(* IEC 61131-3 sources: ia2/library/process-control/pous, 45 files *)

(* ---- fb_alarm_dev.st ---- *)
(*
  FB_ALARM_DEV — deviation alarm (pv over/under deviation from sp), deadband + delay + acknowledge latch.

  ~ Deviation alarm (over/under deviation), standard for loop monitoring.

  Purpose: loop-performance monitoring: alarm on a control deviation that persistently
  exceeds its limit (a stuck valve, an abrupt load change, lost tuning, a failed actuator).
  Behavior (follows the FB_ALARM_HL deadband+delay+latch pattern):
    dev := pv - sp.
    Over deviation:  dev > dev_h sets; dev < dev_h - deadband resets.
    Under deviation: dev < -dev_l sets; dev > -dev_l + deadband resets (dev_l supplied positive).
    Each trips after persisting for delay_s; output = trip OR (latched AND NOT ack)
    -- while the condition exists the alarm stays on, after it clears it is held until acknowledged.

  Inputs:
    pv       REAL  process value
    sp       REAL  setpoint (feed the same sp source as FB_PID; if the PID uses sp_rate,
                   prefer feeding the actual working sp after the ramp)
    dev_h    REAL  over-deviation limit (allowed amount pv may exceed sp)
    dev_l    REAL  under-deviation limit (allowed amount pv may fall below sp, supplied positive)
    deadband REAL  deadband (hysteresis, engineering units)
    delay_s  REAL  alarm delay s (0 = immediate)
    dt_s     REAL  sample period s
    ack      BOOL  acknowledge (level-active)
  Outputs:
    h_alm   BOOL  over-deviation alarm (latched)
    l_alm   BOOL  under-deviation alarm (latched)
    any_alm BOOL  any deviation alarm
*)
FUNCTION_BLOCK FB_ALARM_DEV
  VAR_INPUT
    pv       : REAL;
    sp       : REAL;
    dev_h    : REAL := 10.0;
    dev_l    : REAL := 10.0;
    deadband : REAL := 0.0;
    delay_s  : REAL := 0.0;
    dt_s     : REAL := 0.1;
    ack      : BOOL := FALSE;
  END_VAR
  VAR_OUTPUT
    h_alm   : BOOL;
    l_alm   : BOOL;
    any_alm : BOOL;
  END_VAR
  VAR
    dv     : REAL; (* pv - sp *)
    h_cond : BOOL;
    l_cond : BOOL;
    h_t    : REAL; (* delay accumulator, manual timing in place of TON *)
    l_t    : REAL;
    h_trip : BOOL;
    l_trip : BOOL;
  END_VAR

  dv := pv - sp;

  (* ---- Over deviation ---- *)
  IF dv > dev_h THEN
    h_cond := TRUE;
  ELSIF dv < dev_h - deadband THEN
    h_cond := FALSE;
  END_IF;
  IF h_cond THEN
    h_t := h_t + dt_s;
  ELSE
    h_t := 0.0;
  END_IF;
  h_trip := h_cond AND (h_t >= delay_s);
  h_alm  := h_trip OR (h_alm AND NOT ack);

  (* ---- Under deviation ---- *)
  IF dv < 0.0 - dev_l THEN
    l_cond := TRUE;
  ELSIF dv > 0.0 - dev_l + deadband THEN
    l_cond := FALSE;
  END_IF;
  IF l_cond THEN
    l_t := l_t + dt_s;
  ELSE
    l_t := 0.0;
  END_IF;
  l_trip := l_cond AND (l_t >= delay_s);
  l_alm  := l_trip OR (l_alm AND NOT ack);

  any_alm := h_alm OR l_alm;
END_FUNCTION_BLOCK

(* ---- fb_alarm_hl.st ---- *)
(*
  FB_ALARM_HL — four-level high/low alarm (H/L/HH/LL) with deadband, delay and simplified ISA-18.2 acknowledge latch.

  Purpose: high/low/high-high/low-low alarms for analog values such as level/temperature/pressure.
  Example: a vessel level LT alarm, with HH interlocking the feed shutdown.

  Behavior (same for each level, independently timed):
    1) Raw limit decision (with deadband hysteresis):
       High type: pv > sp sets; pv < sp - deadband resets.
       Low type:  pv < sp sets; pv > sp + deadband resets.
    2) Delay: the limit condition must persist for delay_s before tripping (internally
       timed by manual dt_s accumulation, not a TON instance, for easy offline testing
       and portability).
    3) Latch (simplified ISA-18.2): alarm output = trip condition OR (latched AND NOT ack).
       That is, while the condition exists the alarm stays on; after the condition
       clears it is held until ack acknowledges and clears it.

  Inputs:
    pv        REAL  process value
    h_sp      REAL  high alarm setpoint
    l_sp      REAL  low alarm setpoint
    hh_sp     REAL  high-high alarm setpoint
    ll_sp     REAL  low-low alarm setpoint
    deadband  REAL  deadband (hysteresis, engineering units)
    delay_s   REAL  alarm delay s (0 = immediate)
    dt_s      REAL  sample period s
    ack       BOOL  acknowledge (level-active)
  Outputs:
    h_alm / l_alm / hh_alm / ll_alm  BOOL  latched alarm outputs
    any_alm                          BOOL  any alarm
    h_cond / l_cond / hh_cond / ll_cond BOOL raw limit flags (with deadband, undelayed, unlatched)
*)
FUNCTION_BLOCK FB_ALARM_HL
  VAR_INPUT
    pv       : REAL;
    h_sp     : REAL := 80.0;
    l_sp     : REAL := 20.0;
    hh_sp    : REAL := 90.0;
    ll_sp    : REAL := 10.0;
    deadband : REAL := 0.0;
    delay_s  : REAL := 0.0;
    dt_s     : REAL := 0.1;
    ack      : BOOL := FALSE;
  END_VAR
  VAR_OUTPUT
    h_alm   : BOOL;
    l_alm   : BOOL;
    hh_alm  : BOOL;
    ll_alm  : BOOL;
    any_alm : BOOL;
    h_cond  : BOOL;
    l_cond  : BOOL;
    hh_cond : BOOL;
    ll_cond : BOOL;
  END_VAR
  VAR
    h_t     : REAL; (* per-level delay accumulator, manual timing in place of TON *)
    l_t     : REAL;
    hh_t    : REAL;
    ll_t    : REAL;
    h_trip  : BOOL;
    l_trip  : BOOL;
    hh_trip : BOOL;
    ll_trip : BOOL;
  END_VAR

  (* ---- High alarm H ---- *)
  IF pv > h_sp THEN
    h_cond := TRUE;
  ELSIF pv < h_sp - deadband THEN
    h_cond := FALSE;
  END_IF;
  IF h_cond THEN
    h_t := h_t + dt_s;
  ELSE
    h_t := 0.0;
  END_IF;
  h_trip := h_cond AND (h_t >= delay_s);
  h_alm  := h_trip OR (h_alm AND NOT ack);

  (* ---- Low alarm L ---- *)
  IF pv < l_sp THEN
    l_cond := TRUE;
  ELSIF pv > l_sp + deadband THEN
    l_cond := FALSE;
  END_IF;
  IF l_cond THEN
    l_t := l_t + dt_s;
  ELSE
    l_t := 0.0;
  END_IF;
  l_trip := l_cond AND (l_t >= delay_s);
  l_alm  := l_trip OR (l_alm AND NOT ack);

  (* ---- High-high alarm HH ---- *)
  IF pv > hh_sp THEN
    hh_cond := TRUE;
  ELSIF pv < hh_sp - deadband THEN
    hh_cond := FALSE;
  END_IF;
  IF hh_cond THEN
    hh_t := hh_t + dt_s;
  ELSE
    hh_t := 0.0;
  END_IF;
  hh_trip := hh_cond AND (hh_t >= delay_s);
  hh_alm  := hh_trip OR (hh_alm AND NOT ack);

  (* ---- Low-low alarm LL ---- *)
  IF pv < ll_sp THEN
    ll_cond := TRUE;
  ELSIF pv > ll_sp + deadband THEN
    ll_cond := FALSE;
  END_IF;
  IF ll_cond THEN
    ll_t := ll_t + dt_s;
  ELSE
    ll_t := 0.0;
  END_IF;
  ll_trip := ll_cond AND (ll_t >= delay_s);
  ll_alm  := ll_trip OR (ll_alm AND NOT ack);

  any_alm := h_alm OR l_alm OR hh_alm OR ll_alm;
END_FUNCTION_BLOCK

(* ---- fb_alarm_roc.st ---- *)
(*
  FB_ALARM_ROC — rate-of-change alarm, with derivative filtering, delay and acknowledge latch.

  ~ Rate-of-change alarm, with the derivative denoised by a first-order filter.

  Purpose: monitoring abnormal rates of change such as temperature runaway, abrupt
  pressure change, level collapse (leak/pipe break).
  Behavior:
    Raw derivative raw_roc := (pv - pv_prev) / dt_s;
    roc is raw_roc through an internal PT1 filter (time constant fixed at 3*dt_s,
    settling in about 4 scans) -- a single-scan difference is extremely sensitive to
    quantization/noise and will false-alarm without filtering; for stronger denoising
    put FB_LAG ahead of pv.
    |roc| > roc_limit trips after persisting for delay_s; latched until ack (same as the
    FB_ALARM_HL pattern: while the condition exists the alarm stays on, after it clears
    it is held until acknowledged).
    roc_limit <= 0 -> monitoring disabled (trip condition always FALSE; a latched output
    still needs ack to clear).
    The first scan only aligns pv_prev and does not evaluate the alarm (avoiding a
    spurious startup derivative); dt_s <= 0 -> hold.

  Inputs:
    pv        REAL  process value
    roc_limit REAL  rate-of-change limit |units|/s (bidirectional)
    delay_s   REAL  alarm delay s (0 = immediate)
    dt_s      REAL  sample period s
    ack       BOOL  acknowledge (level-active)
  Outputs:
    alm BOOL  rate-of-change alarm (latched)
    roc REAL  filtered rate of change units/s (signed, usable for trend display)
*)
FUNCTION_BLOCK FB_ALARM_ROC
  VAR_INPUT
    pv        : REAL;
    roc_limit : REAL := 10.0;
    delay_s   : REAL := 0.0;
    dt_s      : REAL := 0.1;
    ack       : BOOL := FALSE;
  END_VAR
  VAR_OUTPUT
    alm : BOOL;
    roc : REAL;
  END_VAR
  VAR
    pv_prev   : REAL;
    raw_roc   : REAL;
    t_f       : REAL; (* derivative filter time constant = 3*dt_s *)
    cond      : BOOL;
    trip      : BOOL;
    alm_t     : REAL; (* delay accumulator *)
    init_done : BOOL;
  END_VAR

  IF dt_s <= 0.0 THEN
    RETURN; (* hold *)
  END_IF;

  IF NOT init_done THEN
    pv_prev := pv; (* first-scan alignment, no alarm evaluation *)
    roc := 0.0;
    init_done := TRUE;
    RETURN;
  END_IF;

  raw_roc := (pv - pv_prev) / dt_s;
  pv_prev := pv;

  (* Internal PT1 denoising: t_f = 3*dt_s fixed (absorbs 1/4 of the new value each scan) *)
  t_f := 3.0 * dt_s;
  roc := roc + dt_s / (t_f + dt_s) * (raw_roc - roc);

  cond := FALSE;
  IF roc_limit > 0.0 THEN
    IF roc > roc_limit OR roc < 0.0 - roc_limit THEN
      cond := TRUE;
    END_IF;
  END_IF;

  IF cond THEN
    alm_t := alm_t + dt_s;
  ELSE
    alm_t := 0.0;
  END_IF;
  trip := cond AND (alm_t >= delay_s);
  alm := trip OR (alm AND NOT ack);
END_FUNCTION_BLOCK

(* ---- fb_alt2.st ---- *)
(*
  FB_ALT2 — dual-valve (dual-device) timed rotator, with two external permissives.

  Purpose: two diverter valves / two pumps rotating on a fixed period for wear balancing.
  Example: dual-permissive diverting with an iron remover + a packing scale:
  permissive1 (iron remover running) or permissive2 (packing scale ready) lost ->
  both valves close at once; after the permissives recover, rotation continues by its
  timer (the rotation selection is held, the timer is cleared and restarts).

  Behavior:
    ok := enable AND permissive1 AND permissive2.
    NOT ok: q1 := FALSE, q2 := FALSE, rotation timer cleared (the selection bit is held,
    and after recovery continues from the last selected channel).
    ok: the timer accumulates by dt_s manually, and at swap_period_s the selection
    switches and the timer clears; q1/q2 output the currently selected channel mutually
    exclusively. swap_period_s <= 0 means no rotation (hold the current channel).

  Inputs:
    enable        BOOL  enable
    swap_period_s REAL  rotation period s
    dt_s          REAL  sample period s
    permissive1   BOOL  external permissive 1 (e.g. iron remover running)
    permissive2   BOOL  external permissive 2 (e.g. packing scale ready)
  Outputs:
    q1 BOOL  valve 1 output
    q2 BOOL  valve 2 output (mutually exclusive with q1; both FALSE when a permissive is lost)
*)
FUNCTION_BLOCK FB_ALT2
  VAR_INPUT
    enable        : BOOL;
    swap_period_s : REAL := 300.0;
    dt_s          : REAL := 0.1;
    permissive1   : BOOL := TRUE;
    permissive2   : BOOL := TRUE;
  END_VAR
  VAR_OUTPUT
    q1 : BOOL;
    q2 : BOOL;
  END_VAR
  VAR
    ok    : BOOL;
    sel2  : BOOL; (* FALSE selects valve 1 / TRUE selects valve 2, held while disabled *)
    run_t : REAL; (* this channel's elapsed run time s, manual timing *)
  END_VAR

  ok := enable AND permissive1 AND permissive2;

  IF NOT ok THEN
    (* Any permissive lost: both valves close, timer cleared, selection held *)
    q1    := FALSE;
    q2    := FALSE;
    run_t := 0.0;
    RETURN;
  END_IF;

  IF dt_s > 0.0 THEN
    run_t := run_t + dt_s;
  END_IF;
  IF swap_period_s > 0.0 AND run_t >= swap_period_s THEN
    run_t := 0.0;
    sel2  := NOT sel2;
  END_IF;

  q1 := NOT sel2;
  q2 := sel2;
END_FUNCTION_BLOCK

(* ---- fb_avg_time.st ---- *)
(*
  FB_AVG_TIME — tumbling-window time average.

  ~ Standard time-average block, the customary form for DCS reporting / steady-quantity monitoring.

  Purpose: full-window averages for reports (e.g. per-minute average flow), noise-robust
  readings of slowly varying quantities, drift monitoring by comparison against the
  instantaneous value.
  Behavior:
    Within the window, sum / count accumulate each scan; avg_run := sum / count is the
    running mean of the current window; when the window is full (accumulated time
    reaches window_s) avg_run is copied into avg, ready is set, and then the
    accumulators are cleared to start the next window (phase subtraction wraps so the
    long-term cadence does not drift).
    While the first window is not yet full, avg temporarily tracks avg_run (to avoid
    outputting 0 at startup) and ready = FALSE flags "not yet a complete-window result";
    after the first window completes ready stays TRUE and avg refreshes only on the
    window-full scan.
    reset level-active: clears the accumulators and ready, restarting the window.
    window_s <= 0 -> pass-through (avg := avg_run := u, ready := TRUE);
    dt_s <= 0 -> hold (no action).
    Note: this block is a tumbling window (one value per window), not a sliding window
    -- a true sliding window needs an array buffer (in this dialect an FB-scope array
    cannot be codegen'd, see README gotcha 7); for continuous "smoothed every scan"
    output, use FB_LAG exponential smoothing as an approximation.

  Inputs:
    u        REAL  input
    window_s REAL  averaging window length s (<= 0 pass-through)
    dt_s     REAL  sample period s
    reset    BOOL  reset (level-active: clear the window and restart)
  Outputs:
    avg     REAL  average of the previous complete window (tracks avg_run while the first window is incomplete)
    avg_run REAL  running mean of the current window
    ready   BOOL  first complete window has finished (avg is trustworthy)
*)
FUNCTION_BLOCK FB_AVG_TIME
  VAR_INPUT
    u        : REAL;
    window_s : REAL := 60.0;
    dt_s     : REAL := 0.1;
    reset    : BOOL := FALSE;
  END_VAR
  VAR_OUTPUT
    avg     : REAL;
    avg_run : REAL;
    ready   : BOOL;
  END_VAR
  VAR
    sum       : REAL; (* current-window accumulated sum *)
    count     : REAL; (* current-window sample count *)
    elapsed_s : REAL; (* current-window accumulated time, manual timing *)
  END_VAR

  IF reset THEN
    sum := 0.0;
    count := 0.0;
    elapsed_s := 0.0;
    avg := 0.0;
    avg_run := 0.0;
    ready := FALSE;
    RETURN;
  END_IF;

  IF window_s <= 0.0 THEN
    avg := u; (* invalid window length: pass-through *)
    avg_run := u;
    ready := TRUE;
    RETURN;
  END_IF;

  IF dt_s <= 0.0 THEN
    RETURN; (* invalid sample period: hold *)
  END_IF;

  sum := sum + u;
  count := count + 1.0;
  elapsed_s := elapsed_s + dt_s;
  avg_run := sum / count;

  IF elapsed_s >= window_s THEN
    (* Window full: copy the result, clear to start the next window (subtraction wrap keeps the long-term cadence) *)
    avg := avg_run;
    ready := TRUE;
    sum := 0.0;
    count := 0.0;
    elapsed_s := elapsed_s - window_s;
  ELSIF NOT ready THEN
    avg := avg_run; (* first window not yet full: avg tracks the running mean to avoid outputting 0 at startup *)
  END_IF;
END_FUNCTION_BLOCK

(* ---- fb_cascade.st ---- *)
(*
  FB_CASCADE — cascade coupling glue (master output -> slave SP mapping + non-cascade tracking back-calculation).

  ~ Standard cascade-coupling block (cascade SP coupling / master tracking
  back-calculation), the customary glue for cascade-loop configuration: only this one
  block sits between the two PIDs.

  Purpose: cascade-loop configuration (temperature master -> flow slave, and the like),
  mapping the master output 0..100% to the slave SP engineering span, and supplying the
  master a tracking value when not in cascade so that putting CAS into/out of service is
  bumpless.
  Behavior:
    CAS (cas_on = TRUE):
      slave_sp := sp_min + master_out / 100 * (sp_max - sp_min)
      master_track := FALSE (the master controls normally).
    Non-CAS:
      slave_sp := slave_sp_local (the operator's local SP given directly to the slave loop);
      master_track := TRUE, master_track_value :=
        (slave_sp_now - sp_min) / (sp_max - sp_min) * 100, clamped 0..100
      -- the master output is forced to "the equivalent percentage of the current slave
      SP", so on the scan that switches back to CAS slave_sp does not jump (bumpless transfer).
      Span not configured (|sp_max - sp_min| < 1E-6) -> tracking value takes 0 (divide-by-zero guard).
    The tracking value is computed every scan (independent of mode), so it is valid the
    instant CAS is removed.
    Pure combinational logic, no internal state.

  Wiring (cascading two FB_PID instances; slave_sp_now is fed the previous scan's working SP):
    casc(master_out := pid_master.out, cas_on := cas_enable,
         sp_min := 0.0, sp_max := 2000.0,
         slave_sp_local := op_sp, slave_sp_now := slave_sp_used);
    slave_sp_used := casc.slave_sp;
    pid_master(pv := temp_pv, sp := temp_sp, ..., dt_s := scan_s,
               track := casc.master_track,
               track_value := casc.master_track_value);
    pid_slave(pv := flow_pv, sp := slave_sp_used, ..., dt_s := scan_s);

  Inputs:
    master_out     REAL  master output 0..100 %
    cas_on         BOOL  cascade enabled (FALSE = slave uses local SP, master tracks)
    sp_min         REAL  slave SP span low (engineering units)
    sp_max         REAL  slave SP span high
    slave_sp_local REAL  slave-loop local SP when not in cascade
    slave_sp_now   REAL  slave-loop current working SP (feed the previous scan's slave_sp, for the tracking back-calculation)
  Outputs:
    slave_sp           REAL  slave-loop setpoint (to pid_slave.sp)
    master_track       BOOL  master tracking command (to pid_master.track)
    master_track_value REAL  master tracking value 0..100 % (to pid_master.track_value)
*)
FUNCTION_BLOCK FB_CASCADE
  VAR_INPUT
    master_out     : REAL;
    cas_on         : BOOL := FALSE;
    sp_min         : REAL := 0.0;
    sp_max         : REAL := 100.0;
    slave_sp_local : REAL := 0.0;
    slave_sp_now   : REAL := 0.0;
  END_VAR
  VAR_OUTPUT
    slave_sp           : REAL;
    master_track       : BOOL;
    master_track_value : REAL;
  END_VAR
  VAR
    span : REAL; (* slave-loop SP span width *)
  END_VAR

  span := sp_max - sp_min;

  (* Tracking value computed every scan: the equivalent percentage of the current slave SP (span not configured -> 0, divide-by-zero guard) *)
  IF (span < 0.000001) AND (span > -0.000001) THEN
    master_track_value := 0.0;
  ELSE
    master_track_value := (slave_sp_now - sp_min) / span * 100.0;
    IF master_track_value < 0.0 THEN
      master_track_value := 0.0;
    ELSIF master_track_value > 100.0 THEN
      master_track_value := 100.0;
    END_IF;
  END_IF;

  IF cas_on THEN
    slave_sp := sp_min + master_out / 100.0 * span;
    master_track := FALSE;
  ELSE
    slave_sp := slave_sp_local;
    master_track := TRUE;
  END_IF;
END_FUNCTION_BLOCK

(* ---- fb_char.st ---- *)
(*
  FB_CHAR — piecewise-linear signal characterization (linear interpolation, up to 8 points).

  ~ Piecewise-linear characterizer, the customary block for valve-characteristic linearization / nonlinear sensors.

  Purpose: valve-characteristic linearization (equal-percentage valve-opening
  compensation), nonlinear sensor calibration, level-to-volume conversion, and any
  monotonic piecewise-linear transform.

  Behavior:
    Take the first n points (x1,y1)..(xn,yn) (n clamped to 2..8); interpolate
    linearly when u falls in segment (xk, xk+1]; u <= x1 -> out := y1; u >= xn ->
    out := yn (clamped at both ends).
    Convention: x must be ascending (no hard check here; a degenerate non-ascending
    segment yields the right-end y).
    In this dialect an ARRAY in FUNCTION_BLOCK scope cannot be codegen'd (see the
    README dialect gotchas), so scalar point pairs x1..x8 / y1..y8 + n are used.

  Inputs:
    u          REAL  input
    n          INT   number of points in use 2..8 (auto-clamped)
    x1..x8     REAL  breakpoint x coordinates (ascending)
    y1..y8     REAL  breakpoint y coordinates
  Outputs:
    out        REAL  characterized output (clamped at both ends)
*)
FUNCTION_BLOCK FB_CHAR
  VAR_INPUT
    u  : REAL;
    n  : INT := 2;
    x1 : REAL := 0.0;
    y1 : REAL := 0.0;
    x2 : REAL := 100.0;
    y2 : REAL := 100.0;
    x3 : REAL := 0.0;
    y3 : REAL := 0.0;
    x4 : REAL := 0.0;
    y4 : REAL := 0.0;
    x5 : REAL := 0.0;
    y5 : REAL := 0.0;
    x6 : REAL := 0.0;
    y6 : REAL := 0.0;
    x7 : REAL := 0.0;
    y7 : REAL := 0.0;
    x8 : REAL := 0.0;
    y8 : REAL := 0.0;
  END_VAR
  VAR_OUTPUT
    out : REAL;
  END_VAR
  VAR
    nn    : INT;  (* clamped point count *)
    xa    : REAL; (* selected segment left end *)
    ya    : REAL;
    xb    : REAL; (* selected segment right end *)
    yb    : REAL;
    span  : REAL;
    found : BOOL;
  END_VAR

  nn := n;
  IF nn < 2 THEN
    nn := 2;
  ELSIF nn > 8 THEN
    nn := 8;
  END_IF;

  (* Low-end clamp *)
  IF u <= x1 THEN
    out := y1;
    RETURN;
  END_IF;

  (* Segment search: take the segment u falls into, (xk, xk+1]; only the first nn points are considered *)
  found := FALSE;
  IF u <= x2 THEN
    xa := x1; ya := y1; xb := x2; yb := y2; found := TRUE;
  ELSIF nn >= 3 AND u <= x3 THEN
    xa := x2; ya := y2; xb := x3; yb := y3; found := TRUE;
  ELSIF nn >= 4 AND u <= x4 THEN
    xa := x3; ya := y3; xb := x4; yb := y4; found := TRUE;
  ELSIF nn >= 5 AND u <= x5 THEN
    xa := x4; ya := y4; xb := x5; yb := y5; found := TRUE;
  ELSIF nn >= 6 AND u <= x6 THEN
    xa := x5; ya := y5; xb := x6; yb := y6; found := TRUE;
  ELSIF nn >= 7 AND u <= x7 THEN
    xa := x6; ya := y6; xb := x7; yb := y7; found := TRUE;
  ELSIF nn >= 8 AND u <= x8 THEN
    xa := x7; ya := y7; xb := x8; yb := y8; found := TRUE;
  END_IF;

  IF found THEN
    span := xb - xa;
    IF span > 0.0 THEN
      out := ya + (u - xa) * (yb - ya) / span;
    ELSE
      out := yb; (* degenerate segment (x not ascending): take the right end *)
    END_IF;
    RETURN;
  END_IF;

  (* High-end clamp: u greater than the nn-th point *)
  CASE nn OF
    3:
      out := y3;
    4:
      out := y4;
    5:
      out := y5;
    6:
      out := y6;
    7:
      out := y7;
    8:
      out := y8;
  ELSE
    out := y2;
  END_CASE;
END_FUNCTION_BLOCK

(* ---- fb_deadtime8.st ---- *)
(*
  FB_DEADTIME8 — dead time / transport delay, 8 scalar taps + linear interpolation.

  ~ Standard dead-time block (dead time / PTt / transport delay), the customary block
  for plant simulation and feedforward dynamic compensation (Smith-predictor-type structures).

  Purpose: plant simulation (in series with FB_LAG it forms a first-order-lag-plus-dead-time
  FOPDT plant), transport-delay matching in a feedforward path, time alignment of
  belt/pipe-conveying measurements.
  Behavior:
    Tap chain z1..z8 (z1 newest, z8 oldest), sampling interval = t_delay_s / 8:
    the phase phase_s accumulates by dt_s manually, and each time a sampling interval
    elapses the whole chain shifts once (z8<-z7<-...<-z1<-u); at most 8 shifts per scan
    (after 8 the whole chain has been filled by u, so the WHILE is bounded and
    scan-deterministic).
    The output interpolates linearly between the two oldest taps by the phase fraction:
      out := z8 + (z7 - z8) * phase_s / period_s
    -- a step input is traversed as a ramp over one sampling interval, so the output is
       continuous with no steps.
    Resolution = t_delay_s / 8: 8 taps is the compromise in an array-free dialect; the
    staircase/interpolation error of the delay time is about 1/8 of the delay --
    adequate for loop tuning; for finer resolution, put two of these blocks in series
    (each carrying half the delay).
    t_delay_s <= 0 -> pass-through (out := u), and the taps fill with u -- when the
    delay is put into service online it starts smoothly from the current value (bumpless).
    reset / first scan: all taps filled with u, out := u, phase cleared.
    dt_s <= 0 -> hold (no action).

  Inputs:
    u         REAL  input
    t_delay_s REAL  dead time s (<= 0 pass-through; changeable online, advances at the new interval)
    dt_s      REAL  sample period s
    reset     BOOL  reset (level-active: taps filled with u, output follows u)
  Outputs:
    out REAL  delayed output (linearly interpolated, continuous)
*)
FUNCTION_BLOCK FB_DEADTIME8
  VAR_INPUT
    u         : REAL;
    t_delay_s : REAL := 0.0;
    dt_s      : REAL := 0.1;
    reset     : BOOL := FALSE;
  END_VAR
  VAR_OUTPUT
    out : REAL;
  END_VAR
  VAR
    z1        : REAL; (* tap chain: z1 newest ... z8 oldest (scalar form for the array-free dialect) *)
    z2        : REAL;
    z3        : REAL;
    z4        : REAL;
    z5        : REAL;
    z6        : REAL;
    z7        : REAL;
    z8        : REAL;
    phase_s   : REAL; (* phase within the current sampling interval, manual timing *)
    period_s  : REAL; (* sampling interval = t_delay_s / 8 *)
    shifts    : REAL; (* shift count this scan (capped at 8: chain already saturated) *)
    init_done : BOOL; (* first-scan alignment flag *)
  END_VAR

  IF reset OR NOT init_done THEN
    z1 := u;
    z2 := u;
    z3 := u;
    z4 := u;
    z5 := u;
    z6 := u;
    z7 := u;
    z8 := u;
    phase_s := 0.0;
    out := u;
    init_done := TRUE;
    RETURN;
  END_IF;

  IF t_delay_s <= 0.0 THEN
    (* Pass-through; taps fill with u, so when the delay is put into service online it starts bumplessly from the current value *)
    z1 := u;
    z2 := u;
    z3 := u;
    z4 := u;
    z5 := u;
    z6 := u;
    z7 := u;
    z8 := u;
    phase_s := 0.0;
    out := u;
    RETURN;
  END_IF;

  IF dt_s <= 0.0 THEN
    RETURN; (* invalid sample period: hold *)
  END_IF;

  period_s := t_delay_s / 8.0;
  phase_s := phase_s + dt_s;

  (* Shift the whole chain once per elapsed sampling interval; capped at 8/scan (when
     dt_s spans several intervals, catch up; after 8 the chain is full of u and further
     shifts are meaningless) -- the WHILE is bounded *)
  shifts := 0.0;
  WHILE (phase_s >= period_s) AND (shifts < 8.0) DO
    z8 := z7;
    z7 := z6;
    z6 := z5;
    z5 := z4;
    z4 := z3;
    z3 := z2;
    z2 := z1;
    z1 := u;
    phase_s := phase_s - period_s;
    shifts := shifts + 1.0;
  END_WHILE;
  IF phase_s >= period_s THEN
    phase_s := 0.0; (* degenerate case dt_s >= t_delay_s: chain is already u, clear phase to prevent accumulation *)
  END_IF;

  (* Interpolate between the two oldest taps by phase fraction: at the shift instant frac=0 -> out=z8(old z7), continuous *)
  out := z8 + (z7 - z8) * phase_s / period_s;
END_FUNCTION_BLOCK

(* ---- fb_debounce.st ---- *)
(*
  FB_DEBOUNCE — discrete-input debounce (independent bidirectional confirmation delay).

  ~ Discrete-input debounce (on/off dual delay), standard for DI processing.

  Purpose: confirming chattering signals such as float level switches, limit switches,
  relay/contactor auxiliary contacts; can also debounce the run_fb/fault inputs of
  FB_DUTY2.
  Behavior:
    u continuously TRUE for t_on_s -> q := TRUE; u continuously FALSE for t_off_s ->
    q := FALSE; any reverse transition in between clears that direction's timer (restart).
    t = 0 means that direction takes effect immediately. The actual confirmation time
    rounds up to a dt_s scan.
    (Manual dt_s accumulation, equivalent to a TON on-confirm + off-confirm, offline-testable.)

  Inputs:
    u       BOOL  raw discrete input
    t_on_s  REAL  set confirmation time s (0 = immediate)
    t_off_s REAL  reset confirmation time s (0 = immediate)
    dt_s    REAL  sample period s
  Outputs:
    q       BOOL  debounced discrete output
*)
FUNCTION_BLOCK FB_DEBOUNCE
  VAR_INPUT
    u       : BOOL;
    t_on_s  : REAL := 0.1;
    t_off_s : REAL := 0.1;
    dt_s    : REAL := 0.1;
  END_VAR
  VAR_OUTPUT
    q : BOOL;
  END_VAR
  VAR
    on_t  : REAL; (* set-direction accumulator *)
    off_t : REAL; (* reset-direction accumulator *)
  END_VAR

  IF u THEN
    off_t := 0.0;
    IF NOT q THEN
      on_t := on_t + dt_s;
      IF on_t >= t_on_s THEN
        q := TRUE;
      END_IF;
    END_IF;
  ELSE
    on_t := 0.0;
    IF q THEN
      off_t := off_t + dt_s;
      IF off_t >= t_off_s THEN
        q := FALSE;
      END_IF;
    END_IF;
  END_IF;
END_FUNCTION_BLOCK

(* ---- fb_deriv.st ---- *)
(*
  FB_DERIV — filtered derivative (du/dt, filter first then difference).

  ~ Standard filtered-derivative block, a staple of every major platform's standard library.

  Purpose: quantifying trend (degC/s, %/s for display/feedforward/custom logic),
  derivative shaping in a feedforward path. Whenever you want "alarm on limit", use
  FB_ALARM_ROC directly (the same filter-difference core + delay/latch).
  Behavior:
    u first passes through an internal PT1 filter (time constant t_filt_s; <= 0 takes
    3*dt_s automatically, settling in about 4 scans), then a backward difference of
    the filtered value:
      u_f := u_f + dt_s / (t_f + dt_s) * (u - u_f)
      out := (u_f - u_f_prev) / dt_s
    A single-scan difference is extremely sensitive to quantization/noise and must be
    filtered, or the output is all spikes -- for stronger noise rejection, increase
    t_filt_s or put FB_LAG ahead of u.
    reset / first scan: the filter state aligns to u, out := 0 (no spurious startup derivative).
    dt_s <= 0 -> hold (no action).

  Inputs:
    u        REAL  input
    t_filt_s REAL  derivative pre-filter time constant s (<= 0 = auto 3*dt_s)
    dt_s     REAL  sample period s
    reset    BOOL  reset/align (level-active: filter state follows u, out cleared)
  Outputs:
    out REAL  filtered rate of change units/s (signed)
*)
FUNCTION_BLOCK FB_DERIV
  VAR_INPUT
    u        : REAL;
    t_filt_s : REAL := 0.0;
    dt_s     : REAL := 0.1;
    reset    : BOOL := FALSE;
  END_VAR
  VAR_OUTPUT
    out : REAL;
  END_VAR
  VAR
    u_f       : REAL; (* PT1-filtered input *)
    u_f_prev  : REAL; (* previous-scan filtered value, for the backward difference *)
    t_f       : REAL; (* filter time constant actually used *)
    init_done : BOOL; (* first-scan alignment flag *)
  END_VAR

  IF dt_s <= 0.0 THEN
    RETURN; (* invalid sample period: hold *)
  END_IF;

  IF reset OR NOT init_done THEN
    u_f := u; (* align the filter state, no spurious startup derivative *)
    u_f_prev := u;
    out := 0.0;
    init_done := TRUE;
    RETURN;
  END_IF;

  t_f := t_filt_s;
  IF t_f <= 0.0 THEN
    t_f := 3.0 * dt_s; (* auto: the minimum noise rejection that settles in about 4 scans *)
  END_IF;

  u_f := u_f + dt_s / (t_f + dt_s) * (u - u_f);
  out := (u_f - u_f_prev) / dt_s;
  u_f_prev := u_f;
END_FUNCTION_BLOCK

(* ---- fb_dose.st ---- *)
(*
  FB_DOSE — batch dosing / batch feeding (coarse/fine two stages + in-flight compensation).

  ~ Standard dosing block (dosing / batch weighing, coarse-fine two-speed feeding +
  early in-flight cutoff), the customary block for batch-scale / batch-feed control.

  Purpose: dosing material from a silo into a weigh hopper / reactor: coarse feed
  approaches the target quickly, fine feed trims, the fine valve closes early by the
  in-flight amount (the material still in flight after the valve closes), and after
  settling the completion and overshoot are reported. The flow input may come from a
  weight derivative or a flowmeter.

  Behavior:
    start rising edge (when idle, not complete, and abort not pressed) begins a new
    batch: qty cleared, enter the feed stage. During feeding/settling, accumulate
    qty := qty + flow * dt_s (flow <= 0 not counted, one of the criteria for material
    fully landed).
      Coarse stage: qty < target - fine_qty -> q_coarse = TRUE (both coarse and fine valves open);
      Fine stage: qty < target - inflight -> q_fine = TRUE; at the point, close the fine
      valve (the in-flight reserve inflight is the in-flight amount held back) and enter
      the settling stage.
      Settling stage: wait for flow <= 0 or a fixed 2 s (whichever first) -> done := TRUE,
      overshoot := qty - target (the actual overshoot once the in-flight material has landed).
    abort level-active: stop both valves immediately, exit feeding/settling, qty
    retained (for stocktaking), done not set.
    After done, start has no effect; reset (level-active) is required to clear
    qty/done/overshoot and begin the next batch.
    Assumes fine_qty >= inflight >= 0 (coarse valve closes first, fine valve closes after);
    dribble after done is no longer counted into qty.
    dt_s <= 0 -> hold this scan, no action (command edges still remembered).

  Inputs:
    start    BOOL  start (rising edge begins a new batch)
    abort    BOOL  abort (level-active: stop valves, retain quantity)
    flow     REAL  instantaneous flow units/s (weight derivative or flowmeter)
    target   REAL  target quantity (same unit as the flow integral)
    fine_qty REAL  fine-feed-stage quantity (close the coarse valve with this much remaining)
    inflight REAL  in-flight amount (close the fine valve with this much remaining)
    dt_s     REAL  sample period s
    reset    BOOL  batch reset (level-active: clear qty/done/overshoot)
  Outputs:
    q_coarse  BOOL  coarse-feed valve
    q_fine    BOOL  fine-feed valve
    qty       REAL  this batch's accumulated quantity
    done      BOOL  this batch complete (set after settling, held until reset)
    overshoot REAL  actual - target after completion (basis for tuning the in-flight amount)
*)
FUNCTION_BLOCK FB_DOSE
  VAR_INPUT
    start    : BOOL;
    abort    : BOOL;
    flow     : REAL;
    target   : REAL := 100.0;
    fine_qty : REAL := 10.0;
    inflight : REAL := 0.0;
    dt_s     : REAL := 0.1;
    reset    : BOOL;
  END_VAR
  VAR_OUTPUT
    q_coarse  : BOOL;
    q_fine    : BOOL;
    qty       : REAL;
    done      : BOOL;
    overshoot : REAL;
  END_VAR
  VAR
    dosing     : BOOL; (* feed stage (coarse/fine) *)
    settling   : BOOL; (* settling-wait stage *)
    settle_t   : REAL; (* settling timer s *)
    prev_start : BOOL; (* start rising-edge memory *)
  END_VAR

  IF reset THEN
    dosing     := FALSE;
    settling   := FALSE;
    settle_t   := 0.0;
    qty        := 0.0;
    done       := FALSE;
    overshoot  := 0.0;
    q_coarse   := FALSE;
    q_fine     := FALSE;
    prev_start := start;
    RETURN;
  END_IF;

  IF abort THEN
    (* Abort: stop valves and exit the stage, qty retained, done not set *)
    dosing   := FALSE;
    settling := FALSE;
    q_coarse := FALSE;
    q_fine   := FALSE;
  END_IF;

  (* start rising edge, idle and not complete -> begin a new batch *)
  IF start AND NOT prev_start AND NOT abort
     AND NOT dosing AND NOT settling AND NOT done THEN
    dosing    := TRUE;
    qty       := 0.0;
    overshoot := 0.0;
    settle_t  := 0.0;
  END_IF;
  prev_start := start;

  IF dt_s <= 0.0 THEN
    RETURN; (* invalid sample period: hold *)
  END_IF;

  (* Accumulate flow during feeding/settling (negative flow not counted) *)
  IF (dosing OR settling) AND flow > 0.0 THEN
    qty := qty + flow * dt_s;
  END_IF;

  IF dosing THEN
    q_coarse := qty < target - fine_qty;
    q_fine   := qty < target - inflight;
    IF NOT q_fine THEN
      (* At the in-flight reserve point: close the fine valve and enter the settling stage *)
      q_coarse := FALSE;
      dosing   := FALSE;
      settling := TRUE;
      settle_t := 0.0;
    END_IF;
  END_IF;

  IF settling THEN
    settle_t := settle_t + dt_s;
    IF flow <= 0.0 OR settle_t >= 2.0 THEN
      settling  := FALSE;
      done      := TRUE;
      overshoot := qty - target;
    END_IF;
  END_IF;
END_FUNCTION_BLOCK

(* ---- fb_duty2.st ---- *)
(*
  FB_DUTY2 — dual-pump duty/standby rotation control.

  ~ Dual-pump duty/standby rotation: select the duty pump by start sequence or run-hour
  balancing, with immediate takeover on fault.

  Purpose: two pumps in a duty/standby arrangement: select the duty pump by rotating
  each start or by balancing accumulated run hours; on a duty-pump fault the standby
  takes over immediately; on a dual fault both stop.
  Behavior (scan-deterministic: no internal timing, only edge memory):
    A demand rising edge selects this round's duty pump, by priority:
      1) exactly one is already running (run_fb TRUE on one side) -> adopt it as duty
         directly (bumpless takeover, avoiding stopping it to start the standby);
      2) alt_mode = 1 -> the lower accumulated hours is duty (hours_a/b fed from two FB_RUNTIME);
      3) alt_mode = 0 (default) -> toggle from the current duty position (including the
         state after a fault takeover, giving natural wear balancing).
    While demand persists: a duty-pump fault with the other healthy -> duty switches
    immediately (takeover); a commanded pump that faults gets no command; a dual fault
    -> both cmd FALSE (the duty selection is held).
    demand withdrawn -> both cmd FALSE.
    Wiring suggestion: feed fault_x from FB_MOTOR's fault or the electrical protection
    relay; feed run_fb_x from the run feedback (debounce a chattering contact with
    FB_DEBOUNCE); leave feedback-timeout fault decision to FB_MOTOR, this block does not
    duplicate the timing.

  Inputs:
    demand   BOOL  system needs a pump (level)
    alt_mode INT   0 = rotate each start / 1 = run-hour balancing
    run_fb_a BOOL  pump A run feedback
    run_fb_b BOOL  pump B run feedback
    fault_a  BOOL  pump A fault
    fault_b  BOOL  pump B fault
    hours_a  REAL  pump A accumulated hours (used by alt_mode=1, fed from FB_RUNTIME.hours)
    hours_b  REAL  pump B accumulated hours (used by alt_mode=1)
    dt_s     REAL  sample period s (this block does not currently time; kept for a uniform library interface)
  Outputs:
    cmd_a     BOOL  pump A start command
    cmd_b     BOOL  pump B start command
    duty_is_a BOOL  the current duty pump is A
*)
FUNCTION_BLOCK FB_DUTY2
  VAR_INPUT
    demand   : BOOL;
    alt_mode : INT := 0;
    run_fb_a : BOOL := FALSE;
    run_fb_b : BOOL := FALSE;
    fault_a  : BOOL := FALSE;
    fault_b  : BOOL := FALSE;
    hours_a  : REAL := 0.0;
    hours_b  : REAL := 0.0;
    dt_s     : REAL := 0.1;
  END_VAR
  VAR_OUTPUT
    cmd_a     : BOOL;
    cmd_b     : BOOL;
    duty_is_a : BOOL;
  END_VAR
  VAR
    prev_demand : BOOL; (* rising-edge memory *)
    rising      : BOOL;
  END_VAR

  rising := demand AND NOT prev_demand;
  prev_demand := demand;

  IF rising THEN
    IF run_fb_a AND NOT run_fb_b THEN
      duty_is_a := TRUE;  (* the already-running pump becomes duty directly, bumpless takeover *)
    ELSIF run_fb_b AND NOT run_fb_a THEN
      duty_is_a := FALSE;
    ELSIF alt_mode = 1 THEN
      duty_is_a := hours_a <= hours_b; (* hour balancing: the lower is duty *)
    ELSE
      duty_is_a := NOT duty_is_a; (* rotate each start (initial FALSE -> first start selects A) *)
    END_IF;
  END_IF;

  IF demand THEN
    (* Fault takeover: duty faults and the other is healthy -> duty switches immediately *)
    IF duty_is_a AND fault_a AND NOT fault_b THEN
      duty_is_a := FALSE;
    ELSIF NOT duty_is_a AND fault_b AND NOT fault_a THEN
      duty_is_a := TRUE;
    END_IF;
    cmd_a := duty_is_a AND NOT fault_a;
    cmd_b := NOT duty_is_a AND NOT fault_b;
  ELSE
    cmd_a := FALSE;
    cmd_b := FALSE;
  END_IF;
END_FUNCTION_BLOCK

(* ---- fb_flow_comp.st ---- *)
(*
  FB_FLOW_COMP — gas-flow pressure/temperature compensation (ideal-gas approximation).

  ~ Standard pressure/temperature compensation block for gas flow, the customary
  block for correcting gas flow to standard / design conditions.

  Purpose: correct gas flow to reference (design) conditions using operating
  pressure/temperature: reading correction for a DP flowmeter calibrated at design
  conditions when operation departs from the design point, and correction of
  volumetric flow to standard conditions. Compensation ratio:
    ratio := (p_abs / p_ref) * (t_ref_k / t_k)   -- density ratio (ideal gas)
    p_abs := p_gauge_kpa + atm_kpa (gauge -> absolute)
    t_k   := t_c + 273.15
  Behavior (mode selects the flowmeter type):
    mode = 0 (square-root DP flowmeter, the flow signal after DP square-root extraction):
      q_comp := q_raw * SQRT(ratio)
      -- DP flow is proportional to SQRT(density), so a density departure from the
         design value is corrected via the square root.
    mode = 1 (linear volumetric, operating volumetric flow corrected to reference conditions):
      q_comp := q_raw * ratio
    Guard: t_k <= 0, t_ref_k <= 0, p_ref_kpa_abs <= 0 or p_abs <= 0
    (invalid measurement/configuration) -> q_comp := q_raw pass-through.
    Pure combinational logic, no internal state.
    Scope note: ideal-gas approximation (no compressibility-factor or humidity
    correction); custody-transfer-grade full-specification energy-metering standard
    algorithms are outside this block's scope.
    Reference conditions default to p_ref = 201.325 kPa(a) (i.e. 100 kPa gauge +
    standard atmosphere), t_ref = 20 degC -- set per the flowmeter design datasheet.

  Inputs:
    q_raw         REAL  raw flow (operating reading)
    p_gauge_kpa   REAL  operating gauge pressure kPa(g)
    t_c           REAL  operating temperature degC
    p_ref_kpa_abs REAL  reference absolute pressure kPa(a) (design condition)
    t_ref_c       REAL  reference temperature degC (design condition)
    atm_kpa       REAL  local atmospheric pressure kPa (gauge -> absolute conversion)
    mode          REAL  0 = square-root DP (multiply by SQRT(ratio)) /
                        1 = linear volumetric (multiply by ratio)
  Outputs:
    q_comp REAL  compensated flow
*)
FUNCTION_BLOCK FB_FLOW_COMP
  VAR_INPUT
    q_raw         : REAL;
    p_gauge_kpa   : REAL;
    t_c           : REAL;
    p_ref_kpa_abs : REAL := 201.325;
    t_ref_c       : REAL := 20.0;
    atm_kpa       : REAL := 101.325;
    mode          : REAL := 0.0;
  END_VAR
  VAR_OUTPUT
    q_comp : REAL;
  END_VAR
  VAR
    p_abs_kpa : REAL; (* operating absolute pressure *)
    t_k       : REAL; (* operating absolute temperature K *)
    t_ref_k   : REAL; (* reference absolute temperature K *)
    ratio     : REAL; (* density ratio (ideal gas) *)
  END_VAR

  p_abs_kpa := p_gauge_kpa + atm_kpa;
  t_k := t_c + 273.15;
  t_ref_k := t_ref_c + 273.15;

  IF (t_k <= 0.0) OR (t_ref_k <= 0.0)
     OR (p_ref_kpa_abs <= 0.0) OR (p_abs_kpa <= 0.0) THEN
    q_comp := q_raw; (* invalid measurement/configuration: pass-through *)
    RETURN;
  END_IF;

  ratio := (p_abs_kpa / p_ref_kpa_abs) * (t_ref_k / t_k);

  IF mode >= 0.5 THEN
    q_comp := q_raw * ratio;       (* 1 = linear volumetric *)
  ELSE
    q_comp := q_raw * SQRT(ratio); (* 0 = square-root DP *)
  END_IF;
END_FUNCTION_BLOCK

(* ---- fb_gain_sched3.st ---- *)
(*
  FB_GAIN_SCHED3 — three-zone gain scheduling (gain scheduling, hysteresis zoning +
  optional zone-boundary linear transition).

  ~ Standard gain scheduler / parameter scheduler (switches the PID parameter set by
  zone of an operating variable), the customary block for segmented tuning of a
  nonlinear plant.

  Purpose: when the plant gain varies greatly with operating point (load segments,
  valve-characteristic segments, the strongly nonlinear pH segment), output a kp/ti/td
  parameter set in three zones of a scheduling variable (load / opening / the PV itself);
  the output feeds the parameter inputs of FB_PID / FB_PID_POS directly -- an online
  parameter change takes effect immediately (both blocks compute their increment/terms
  from the current parameters).

  Behavior:
    Zoning (u_sched against the two boundaries x12 / x23, assuming x12 < x23):
      zone 1: u <= x12; zone 2: x12 < u <= x23; zone 3: u > x23.
    Hysteresis: a zone change requires crossing the boundary +/- hyst (preventing
    chatter near a boundary from toggling parameters back and forth); the first scan
    seeds by plain comparison. A large step can jump two zones within one scan (it
    settles by stepwise migration).
    Parameter output:
      interp = FALSE: take the current zone's parameter set (hysteresis switching, with
      stepped parameters -- feeding incremental FB_PID is naturally bumpless, feeding
      FB_PID_POS recomputes the P term immediately at the new kp);
      interp = TRUE and hyst > 0: when u falls within +/-hyst of a boundary the two
      zones' parameters transition linearly (parameter output continuous, determined by
      u_sched alone; zone still gives its discrete indication by hysteresis).
    Note: when interp mixes a zone with ti = 0 (integral off) and one with ti > 0, the
    transition segment produces a very small ti (very strong integral) -- each zone's
    ti/td should be all 0 or all non-zero.

  Inputs:
    u_sched         REAL  scheduling variable (load / valve position / PV, etc.)
    x12             REAL  zone 1/2 boundary
    x23             REAL  zone 2/3 boundary (> x12, and the two transition bands must not overlap)
    hyst            REAL  zone-boundary hysteresis half-width (0 = no hysteresis)
    interp          BOOL  TRUE = linear parameter transition within +/-hyst of a boundary
    kp1, ti1_s, td1_s REAL  zone 1 parameter set
    kp2, ti2_s, td2_s REAL  zone 2 parameter set
    kp3, ti3_s, td3_s REAL  zone 3 parameter set
  Outputs:
    kp_out   REAL  scheduled proportional gain (to the PID's kp)
    ti_out_s REAL  scheduled integral time s
    td_out_s REAL  scheduled derivative time s
    zone     REAL  current zone 1 / 2 / 3 (hysteresis decision)
*)
FUNCTION_BLOCK FB_GAIN_SCHED3
  VAR_INPUT
    u_sched : REAL;
    x12     : REAL := 33.3;
    x23     : REAL := 66.6;
    hyst    : REAL := 0.0;
    interp  : BOOL := FALSE;
    kp1     : REAL := 1.0;
    ti1_s   : REAL := 0.0;
    td1_s   : REAL := 0.0;
    kp2     : REAL := 1.0;
    ti2_s   : REAL := 0.0;
    td2_s   : REAL := 0.0;
    kp3     : REAL := 1.0;
    ti3_s   : REAL := 0.0;
    td3_s   : REAL := 0.0;
  END_VAR
  VAR_OUTPUT
    kp_out   : REAL;
    ti_out_s : REAL;
    td_out_s : REAL;
    zone     : REAL;
  END_VAR
  VAR
    f : REAL; (* interpolation fraction within the transition band 0..1 *)
  END_VAR

  (* 1) Zone selection (hysteresis): first scan zone = 0 -> seed by plain comparison *)
  IF zone < 0.5 THEN
    IF u_sched <= x12 THEN
      zone := 1.0;
    ELSIF u_sched <= x23 THEN
      zone := 2.0;
    ELSE
      zone := 3.0;
    END_IF;
  END_IF;

  (* Stepwise migration (test 1->2, 3->2 first, then 2->1/2->3: a large step settles in one scan) *)
  IF zone <= 1.5 THEN
    IF u_sched > x12 + hyst THEN
      zone := 2.0;
    END_IF;
  END_IF;
  IF zone >= 2.5 THEN
    IF u_sched < x23 - hyst THEN
      zone := 2.0;
    END_IF;
  END_IF;
  IF zone >= 1.5 AND zone <= 2.5 THEN
    IF u_sched > x23 + hyst THEN
      zone := 3.0;
    ELSIF u_sched < x12 - hyst THEN
      zone := 1.0;
    END_IF;
  END_IF;

  (* 2) Zone parameters (discrete values, hysteresis switching) *)
  IF zone <= 1.5 THEN
    kp_out   := kp1;
    ti_out_s := ti1_s;
    td_out_s := td1_s;
  ELSIF zone <= 2.5 THEN
    kp_out   := kp2;
    ti_out_s := ti2_s;
    td_out_s := td2_s;
  ELSE
    kp_out   := kp3;
    ti_out_s := ti3_s;
    td_out_s := td3_s;
  END_IF;

  (* 3) interp: linear transition within +/-hyst of a boundary (parameters continuous,
        determined by u_sched alone, overriding the discrete values above; the zone
        output is unaffected) *)
  IF interp AND hyst > 0.0 THEN
    IF (u_sched > x12 - hyst) AND (u_sched < x12 + hyst) THEN
      f := (u_sched - (x12 - hyst)) / (2.0 * hyst);
      kp_out   := kp1 + f * (kp2 - kp1);
      ti_out_s := ti1_s + f * (ti2_s - ti1_s);
      td_out_s := td1_s + f * (td2_s - td1_s);
    ELSIF (u_sched > x23 - hyst) AND (u_sched < x23 + hyst) THEN
      f := (u_sched - (x23 - hyst)) / (2.0 * hyst);
      kp_out   := kp2 + f * (kp3 - kp2);
      ti_out_s := ti2_s + f * (ti3_s - ti2_s);
      td_out_s := td2_s + f * (td3_s - td2_s);
    ELSIF u_sched <= x12 - hyst THEN
      kp_out   := kp1;
      ti_out_s := ti1_s;
      td_out_s := td1_s;
    ELSIF u_sched >= x23 + hyst THEN
      kp_out   := kp3;
      ti_out_s := ti3_s;
      td_out_s := td3_s;
    ELSE
      kp_out   := kp2; (* between the two transition bands: pure zone 2 *)
      ti_out_s := ti2_s;
      td_out_s := td2_s;
    END_IF;
  END_IF;
END_FUNCTION_BLOCK

(* ---- fb_hilo_fill.st ---- *)
(*
  FB_HILO_FILL — high-close, low-open tank/silo replenishment control.

  Purpose: below the low setpoint open the supply valve, above the high setpoint close
  it, hold the current state in between (equivalent to a low-side-on hysteresis switch,
  given a dedicated name for readability in configuration).
  Example: circulating-tank make-up: pv <= l_sp opens the make-up valve, pv >= h_sp closes it.

  Behavior:
    pv <= l_sp -> valve_open := TRUE (low-open)
    pv >= h_sp -> valve_open := FALSE (high-close)
    l_sp < pv < h_sp -> hold.
  Assumes l_sp < h_sp; if reversed, the high test takes priority (opens then is
  immediately closed, output FALSE).

  Inputs:
    pv   REAL  level process value
    h_sp REAL  high setpoint (close)
    l_sp REAL  low setpoint (open)
  Outputs:
    valve_open BOOL  supply-valve output (TRUE open)
*)
FUNCTION_BLOCK FB_HILO_FILL
  VAR_INPUT
    pv   : REAL;
    h_sp : REAL := 85.0;
    l_sp : REAL := 15.0;
  END_VAR
  VAR_OUTPUT
    valve_open : BOOL;
  END_VAR

  IF pv >= h_sp THEN
    valve_open := FALSE; (* high-close, priority *)
  ELSIF pv <= l_sp THEN
    valve_open := TRUE;  (* low-open *)
  END_IF;
  (* Hold in between *)
END_FUNCTION_BLOCK

(* ---- fb_hyst.st ---- *)
(*
  FB_HYST — bidirectional hysteresis (deadband) switch.

  Purpose: on/off control of an analog value with hysteresis, avoiding chatter at the threshold.
  Example: current control of a feeder -- current above on_sp stops feeding, below
  off_sp resumes (low-side-on direction); or temperature above on_sp starts a fan, below
  off_sp stops it (high-side-on direction).

  Behavior (direction decided automatically from the setpoints):
    on_sp > off_sp (high-side-on): pv >= on_sp sets; pv <= off_sp resets; holds in between.
    on_sp < off_sp (low-side-on):  pv <= on_sp sets; pv >= off_sp resets; holds in between.
    on_sp = off_sp (degenerate):   out := pv >= on_sp (plain comparator, no hysteresis).

  Inputs:
    pv     REAL  process value
    on_sp  REAL  switch-on setpoint
    off_sp REAL  switch-off setpoint
  Outputs:
    out    BOOL  switch output
*)
FUNCTION_BLOCK FB_HYST
  VAR_INPUT
    pv     : REAL;
    on_sp  : REAL;
    off_sp : REAL;
  END_VAR
  VAR_OUTPUT
    out : BOOL;
  END_VAR

  IF on_sp > off_sp THEN
    (* High-side-on *)
    IF pv >= on_sp THEN
      out := TRUE;
    ELSIF pv <= off_sp THEN
      out := FALSE;
    END_IF;
  ELSIF on_sp < off_sp THEN
    (* Low-side-on *)
    IF pv <= on_sp THEN
      out := TRUE;
    ELSIF pv >= off_sp THEN
      out := FALSE;
    END_IF;
  ELSE
    (* Setpoints equal: degenerate to a plain comparator *)
    out := pv >= on_sp;
  END_IF;
END_FUNCTION_BLOCK

(* ---- fb_integ.st ---- *)
(*
  FB_INTEG — general-purpose integrator (with hold/reset/preset and output clamp).

  ~ Standard integrator block, a staple of every major platform's standard library.

  Purpose: deviation integration (monitoring accumulated quantities such as degC*s),
  simple material/energy totals, the integral element in plant simulation, the
  integral path of a custom control algorithm.
  Difference from FB_TOTALIZER: TOTALIZER is a flow-totalizing block fixed at /3600;
  this block is general integration out := out + k * u * dt_s, with hold/preset/clamp.
  Behavior (command priority reset > preset > hold > integrate):
    reset  level-active: out := 0, limit flags cleared;
    preset level-active: out := preset_value (then clamped as usual);
    hold   level-active: integration paused, output held (clamp and limit flags still refresh);
    otherwise: out := out + k * u * dt_s, clamped to [out_min, out_max].
    q_hi / q_lo indicate the output at the high/low limit (anti-windup: at a limit, a
    reverse input exits immediately).
    dt_s <= 0 -> hold this scan (reset/preset are level commands, not subject to this).

  Inputs:
    u            REAL  integrand input
    k            REAL  integral gain (1/s; dimension defined by the caller)
    dt_s         REAL  sample period s
    hold         BOOL  pause integration (level-active)
    reset        BOOL  reset to 0 (level-active, highest priority)
    preset       BOOL  preset (level-active, takes priority over hold)
    preset_value REAL  preset value
    out_min      REAL  output low limit (default -1.0E38 ~ unlimited)
    out_max      REAL  output high limit (default +1.0E38 ~ unlimited)
  Outputs:
    out  REAL  integral output (clamped)
    q_hi BOOL  at high limit
    q_lo BOOL  at low limit
*)
FUNCTION_BLOCK FB_INTEG
  VAR_INPUT
    u            : REAL;
    k            : REAL := 1.0;
    dt_s         : REAL := 0.1;
    hold         : BOOL := FALSE;
    reset        : BOOL := FALSE;
    preset       : BOOL := FALSE;
    preset_value : REAL := 0.0;
    out_min      : REAL := -1.0E38;
    out_max      : REAL := 1.0E38;
  END_VAR
  VAR_OUTPUT
    out  : REAL;
    q_hi : BOOL;
    q_lo : BOOL;
  END_VAR

  IF reset THEN
    out := 0.0;
    q_hi := FALSE;
    q_lo := FALSE;
    RETURN;
  END_IF;

  IF preset THEN
    out := preset_value; (* after preset, fall through to the clamp below as usual *)
  ELSIF NOT hold THEN
    IF dt_s <= 0.0 THEN
      RETURN; (* invalid sample period: hold *)
    END_IF;
    out := out + k * u * dt_s;
  END_IF;
  (* While hold is active: no integration, just refresh the clamp and limit flags as usual *)

  q_hi := FALSE;
  q_lo := FALSE;
  IF out >= out_max THEN
    out := out_max;
    q_hi := TRUE;
  ELSIF out <= out_min THEN
    out := out_min;
    q_lo := TRUE;
  END_IF;
END_FUNCTION_BLOCK

(* ---- fb_interlock8.st ---- *)
(*
  FB_INTERLOCK8 — 8-channel interlock summary + first-out recording.

  ~ Interlock summary + first-out capture (first-out annunciation, after the ISA-18.1 first-out-window concept).

  Purpose: trip-cause tracing for a unit interlock: summarize multiple conditions into a
  single trip bit and latch the channel that acted first, to locate the trip root cause
  afterward (consequential actions after the first-out do not overwrite the record).
  Behavior:
    Effective condition ax := cx AND enablex (enablex default TRUE; setting FALSE = bypass that channel).
    tripped := any effective condition OR (latched AND NOT reset)
    -- while any condition exists the alarm stays on; after all conditions clear it is
    held until reset (equivalent to "reset AND all clear" to reset; reset has no effect
    while a condition is uncleared).
    First-out capture: the scan where tripped goes FALSE->TRUE records the lowest channel
    number acting at that moment (on a tie, the lowest number). During the interlock hold,
    later actions do not overwrite the first-out; on a successful reset (tripped returns
    FALSE) first_out is cleared to 0.
    cx semantics: TRUE = that condition has acted (trip direction). Invert normally-closed
    signals externally.

  Inputs:
    c1..c8           BOOL  interlock conditions (TRUE = acted/over-limit)
    enable1..enable8 BOOL  per-channel in service (default TRUE; FALSE = bypass)
    reset            BOOL  reset (level-active; effective only after all conditions clear)
  Outputs:
    tripped   BOOL  interlock acted (latched)
    first_out INT   first-out channel number 1..8, 0 = none
*)
FUNCTION_BLOCK FB_INTERLOCK8
  VAR_INPUT
    c1      : BOOL := FALSE;
    c2      : BOOL := FALSE;
    c3      : BOOL := FALSE;
    c4      : BOOL := FALSE;
    c5      : BOOL := FALSE;
    c6      : BOOL := FALSE;
    c7      : BOOL := FALSE;
    c8      : BOOL := FALSE;
    enable1 : BOOL := TRUE;
    enable2 : BOOL := TRUE;
    enable3 : BOOL := TRUE;
    enable4 : BOOL := TRUE;
    enable5 : BOOL := TRUE;
    enable6 : BOOL := TRUE;
    enable7 : BOOL := TRUE;
    enable8 : BOOL := TRUE;
    reset   : BOOL := FALSE;
  END_VAR
  VAR_OUTPUT
    tripped   : BOOL;
    first_out : INT;
  END_VAR
  VAR
    a1    : BOOL; (* effective condition after in-service gating *)
    a2    : BOOL;
    a3    : BOOL;
    a4    : BOOL;
    a5    : BOOL;
    a6    : BOOL;
    a7    : BOOL;
    a8    : BOOL;
    any_c : BOOL;
    was   : BOOL; (* previous-scan tripped, to capture the first-out edge *)
  END_VAR

  a1 := c1 AND enable1;
  a2 := c2 AND enable2;
  a3 := c3 AND enable3;
  a4 := c4 AND enable4;
  a5 := c5 AND enable5;
  a6 := c6 AND enable6;
  a7 := c7 AND enable7;
  a8 := c8 AND enable8;
  any_c := a1 OR a2 OR a3 OR a4 OR a5 OR a6 OR a7 OR a8;

  was := tripped;
  tripped := any_c OR (tripped AND NOT reset);

  IF tripped AND NOT was THEN
    (* New trip event: record the first-out (on a tie, the lowest number) *)
    IF a1 THEN
      first_out := 1;
    ELSIF a2 THEN
      first_out := 2;
    ELSIF a3 THEN
      first_out := 3;
    ELSIF a4 THEN
      first_out := 4;
    ELSIF a5 THEN
      first_out := 5;
    ELSIF a6 THEN
      first_out := 6;
    ELSIF a7 THEN
      first_out := 7;
    ELSIF a8 THEN
      first_out := 8;
    END_IF;
  ELSIF NOT tripped THEN
    first_out := 0; (* successful reset clears the first-out *)
  END_IF;
END_FUNCTION_BLOCK

(* ---- fb_lag.st ---- *)
(*
  FB_LAG — first-order lag filter (PT1 / first-order lag).

  ~ Standard first-order lag filter (PT1 / LAG), a staple of every major platform's standard library.

  Purpose: analog noise rejection, measurement smoothing, pre-filtering ahead of
  derivative / rate-of-change computation.
  Algorithm (backward-Euler discretization, unconditionally stable):
    out := out + dt_s / (t_s + dt_s) * (u - out)
  Notes:
    t_s <= 0 -> pass-through (out := u); dt_s <= 0 -> hold (no action);
    reset level-active -> out := u (filter alignment, bumpless startup);
    the first scan auto-aligns (out := u) to avoid a startup transient
    crawling up from 0.

  Inputs:
    u     REAL  input
    t_s   REAL  filter time constant s (0 = pass-through)
    dt_s  REAL  sample period s
    reset BOOL  reset/align (level-active: out follows u)
  Outputs:
    out   REAL  filtered output
*)
FUNCTION_BLOCK FB_LAG
  VAR_INPUT
    u     : REAL;
    t_s   : REAL := 1.0;
    dt_s  : REAL := 0.1;
    reset : BOOL := FALSE;
  END_VAR
  VAR_OUTPUT
    out : REAL;
  END_VAR
  VAR
    init_done : BOOL; (* first-scan alignment flag *)
  END_VAR

  IF reset OR NOT init_done THEN
    out := u;
    init_done := TRUE;
    RETURN;
  END_IF;

  IF t_s <= 0.0 THEN
    out := u; (* pass-through *)
    RETURN;
  END_IF;

  IF dt_s <= 0.0 THEN
    RETURN; (* invalid sample period: hold *)
  END_IF;

  out := out + dt_s / (t_s + dt_s) * (u - out);
END_FUNCTION_BLOCK

(* ---- fb_leadlag.st ---- *)
(*
  FB_LEADLAG — lead-lag compensator (feedforward-path dynamic shaping).

  ~ Standard lead-lag compensation, the customary block for dynamic shaping of a feedforward path.

  Purpose: dynamic matching for feedforward compensation: pass the feedforward
  signal through (1 + s*lead_s)/(1 + s*lag_s) to compensate the time difference
  between the disturbance path and the control path. lead_s > lag_s leads (speeds
  up the response), lead_s < lag_s lags (buffers). The output typically feeds the
  ff input of FB_PID.

  Discrete approximation (standard decomposition: internal PT1 + pass-through mix):
    filt := filt + dt_s / (lag_s + dt_s) * (u - filt)   -- internal first-order lag
    out  := u * (lead_s / lag_s) + filt * (1 - lead_s / lag_s)
  Compared with the continuous transfer function: steady-state gain 1, high-frequency
  gain lead_s/lag_s (first-order approximation; approaches the continuous solution
  when dt_s << lag_s).
  Notes:
    lag_s <= 0 -> pass-through (out := u, filt follows);
    lead_s = 0 -> degenerates to a pure PT1; lead_s = lag_s -> pass-through;
    when lead_s/lag_s is much greater than 1 the high-frequency gain is large, so
    watch for input-noise amplification;
    reset or first scan -> filt := u, out := u (bumpless startup); dt_s <= 0 -> hold.

  Inputs:
    u      REAL  input
    lead_s REAL  lead time constant s
    lag_s  REAL  lag time constant s (0 = pass-through)
    dt_s   REAL  sample period s
    reset  BOOL  reset/align (level-active)
  Outputs:
    out    REAL  compensated output
*)
FUNCTION_BLOCK FB_LEADLAG
  VAR_INPUT
    u      : REAL;
    lead_s : REAL := 0.0;
    lag_s  : REAL := 1.0;
    dt_s   : REAL := 0.1;
    reset  : BOOL := FALSE;
  END_VAR
  VAR_OUTPUT
    out : REAL;
  END_VAR
  VAR
    filt      : REAL; (* internal PT1 state *)
    gain_hf   : REAL; (* lead_s / lag_s *)
    init_done : BOOL;
  END_VAR

  IF reset OR NOT init_done THEN
    filt := u;
    out := u;
    init_done := TRUE;
    RETURN;
  END_IF;

  IF lag_s <= 0.0 THEN
    filt := u;
    out := u; (* pass-through *)
    RETURN;
  END_IF;

  IF dt_s <= 0.0 THEN
    RETURN; (* hold *)
  END_IF;

  filt := filt + dt_s / (lag_s + dt_s) * (u - filt);
  gain_hf := lead_s / lag_s;
  out := u * gain_hf + filt * (1.0 - gain_hf);
END_FUNCTION_BLOCK

(* ---- fb_limit.st ---- *)
(*
  FB_LIMIT — value limiter (high-low clamp + limit indication).

  ~ Standard limiter (limiter / high-low clamp), a staple of every major platform's standard library.

  Purpose: safe clamping of setpoint/output values, cascade outer-loop output limiting,
  operator-input validation, the last line of protection for a bare downstream actuator.
  Behavior (pure combinational logic, no internal state):
    out := u clamped to [lo, hi]; q_hi / q_lo indicate clamping in progress (u over the high/low limit).
    Configuration error lo > hi -> out := (lo + hi) / 2, with q_hi and q_lo both TRUE
    -- both limit flags lit at once cannot occur physically and serves purely as a
    configuration-error signal, easy for a supervisory alarm to catch.

  Inputs:
    u  REAL  input
    lo REAL  low limit
    hi REAL  high limit (assumes lo <= hi; reversed triggers the configuration-error signal)
  Outputs:
    out  REAL  clamped output
    q_hi BOOL  over high limit (clamping at hi)
    q_lo BOOL  over low limit (clamping at lo; TRUE together with q_hi = lo > hi configuration error)
*)
FUNCTION_BLOCK FB_LIMIT
  VAR_INPUT
    u  : REAL;
    lo : REAL := 0.0;
    hi : REAL := 100.0;
  END_VAR
  VAR_OUTPUT
    out  : REAL;
    q_hi : BOOL;
    q_lo : BOOL;
  END_VAR

  IF lo > hi THEN
    (* Configuration error: output the midpoint, both limit flags lit as the error signal *)
    out := (lo + hi) / 2.0;
    q_hi := TRUE;
    q_lo := TRUE;
    RETURN;
  END_IF;

  IF u > hi THEN
    out := hi;
    q_hi := TRUE;
    q_lo := FALSE;
  ELSIF u < lo THEN
    out := lo;
    q_hi := FALSE;
    q_lo := TRUE;
  ELSE
    out := u;
    q_hi := FALSE;
    q_lo := FALSE;
  END_IF;
END_FUNCTION_BLOCK

(* ---- fb_manstation.st ---- *)
(*
  FB_MANSTATION — manual loader / bias station.

  ~ Standard manual station + bias station (manual station / auto-manual station with
  bias), the standard operating layer between a controller output and an actuator,
  found in every major DCS/PLC standard library.

  Purpose: placed between a controller output and an actuator: in auto it passes through
  (with optional bias and rate limiting); in manual the operator sets the output
  directly; balance guarantees a bumpless manual->auto transfer. It can also serve
  standalone as a pure manual loader (auto := FALSE, always manual) or a pure bias /
  rate-limit station.

  Behavior:
    Auto (auto = TRUE): out approaches (auto_in + bias + corr) --
      when rate > 0 limited to rate units/second, rate = 0 steps directly; clamped to
      [out_min, out_max]. corr is the internal bias correction back-calculated at a balance transfer.
    Manual (auto = FALSE): out := manual_out (clamped, not rate-limited),
      tracking := TRUE.
    Bumpless transfer (balance = TRUE): the manual->auto transition edge back-calculates
      corr := out - auto_in - bias
    -- out is continuous at the transfer instant; afterward changes in auto_in/bias take
    effect as usual, and corr is held until recomputed at the next transfer. When
    balance = FALSE, corr is always 0 (the transfer step is ridden out by the rate
    limit; rate = 0 means a step).
    First scan: out aligns directly to the current mode's target value (no climb from 0).
    dt_s <= 0 -> hold this scan, no action.
    Note: bias is the nominal bias written by the operator/supervisory level; corr is
    the block's self-trimming correction, and the two add. To "clear" the historical
    correction, set balance := FALSE for one scan.

  Inputs:
    auto_in    REAL  auto input (upstream controller output)
    auto       BOOL  TRUE auto / FALSE manual
    manual_out REAL  manual output value
    bias       REAL  bias (added in auto)
    rate       REAL  auto-output rate limit units/s (0 = no rate limit)
    out_min    REAL  output low limit
    out_max    REAL  output high limit
    balance    BOOL  TRUE = back-calculate the bias correction on a manual->auto transfer (bumpless)
    dt_s       REAL  sample period s
  Outputs:
    out      REAL  station output (clamped in every mode)
    tracking BOOL  in manual (the upstream controller can use this bit for output tracking)
*)
FUNCTION_BLOCK FB_MANSTATION
  VAR_INPUT
    auto_in    : REAL;
    auto       : BOOL := TRUE;
    manual_out : REAL := 0.0;
    bias       : REAL := 0.0;
    rate       : REAL := 0.0;
    out_min    : REAL := 0.0;
    out_max    : REAL := 100.0;
    balance    : BOOL := TRUE;
    dt_s       : REAL := 0.1;
  END_VAR
  VAR_OUTPUT
    out      : REAL;
    tracking : BOOL;
  END_VAR
  VAR
    corr      : REAL; (* internal bias correction back-calculated by balance *)
    target    : REAL; (* auto target = auto_in + bias + corr *)
    delta     : REAL;
    step      : REAL;
    prev_auto : BOOL; (* transfer-edge memory *)
    init_done : BOOL; (* first-scan alignment flag *)
  END_VAR

  IF dt_s <= 0.0 THEN
    RETURN; (* invalid sample period: hold *)
  END_IF;

  IF NOT balance THEN
    corr := 0.0;
  END_IF;

  IF NOT init_done THEN
    (* First scan: align directly to the current mode's target, no climb from 0 *)
    IF auto THEN
      out := auto_in + bias;
    ELSE
      out := manual_out;
    END_IF;
    IF out > out_max THEN
      out := out_max;
    ELSIF out < out_min THEN
      out := out_min;
    END_IF;
    tracking := NOT auto;
    prev_auto := auto;
    init_done := TRUE;
    RETURN;
  END_IF;

  (* Manual->auto transition edge: balance back-calculates the correction so out is continuous *)
  IF auto AND NOT prev_auto AND balance THEN
    corr := out - auto_in - bias;
  END_IF;
  prev_auto := auto;

  IF NOT auto THEN
    (* Manual: set directly (clamped, not rate-limited) *)
    out := manual_out;
    IF out > out_max THEN
      out := out_max;
    ELSIF out < out_min THEN
      out := out_min;
    END_IF;
    tracking := TRUE;
    RETURN;
  END_IF;
  tracking := FALSE;

  (* Auto: approach auto_in + bias + corr at the rate limit (rate = 0 steps) *)
  target := auto_in + bias + corr;
  IF rate > 0.0 THEN
    delta := target - out;
    step := rate * dt_s;
    IF delta > step THEN
      out := out + step;
    ELSIF delta < 0.0 - step THEN
      out := out - step;
    ELSE
      out := target;
    END_IF;
  ELSE
    out := target;
  END_IF;

  IF out > out_max THEN
    out := out_max;
  ELSIF out < out_min THEN
    out := out_min;
  END_IF;
END_FUNCTION_BLOCK

(* ---- fb_mid3.st ---- *)
(*
  FB_MID3 — median select / 2oo3 analog voting.

  ~ Standard median-select / redundant-measurement voting block (median selector,
  2oo3 voting), the customary block for redundant-transmitter signal selection.

  Purpose: median of three redundant transmitters (rejects single-point drift/jump),
  average of dual redundancy, bad-value degradation of critical measurements (pair
  with the inverse of FB_SCALE fault as good_x).
  Behavior (degrades by the number of good channels n_good):
    3 good -> take the median (naturally rejects single-channel drift);
    2 good -> take the average of the two good channels;
    1 good -> pass that channel through;
    0 good -> out holds the previous scan's value, q_fail = TRUE (level, not latched).
    Deviation monitor: when dev_max > 0, the difference between any two good channels
    > dev_max -> q_dev (signals that drift between redundant channels has widened and
    a transmitter check is due; dev_max <= 0 disables the monitor).
    good_x takes the bad-value decision (transmitter open-circuit/over-range, e.g. the
    inverse of FB_SCALE.fault), defaulting to TRUE = all good.
    Note: when there are 0 good on the very first scan, out is its initial value 0 (no
    history to hold); the held value during q_fail is "the voted value from the last
    time a good channel existed".

  Inputs:
    a, b, c                REAL  three redundant measurements
    good_a, good_b, good_c BOOL  per-channel validity (default TRUE; FALSE = excluded)
    dev_max                REAL  deviation-monitor limit between good channels (<= 0 = disabled)
  Outputs:
    out    REAL  voted output (held when 0 good)
    n_good REAL  current number of good channels 0..3
    q_dev  BOOL  deviation between good channels over limit
    q_fail BOOL  all channels failed (output is in hold)
*)
FUNCTION_BLOCK FB_MID3
  VAR_INPUT
    a       : REAL;
    b       : REAL;
    c       : REAL;
    good_a  : BOOL := TRUE;
    good_b  : BOOL := TRUE;
    good_c  : BOOL := TRUE;
    dev_max : REAL := 0.0;
  END_VAR
  VAR_OUTPUT
    out    : REAL;
    n_good : REAL;
    q_dev  : BOOL;
    q_fail : BOOL;
  END_VAR

  n_good := 0.0;
  IF good_a THEN
    n_good := n_good + 1.0;
  END_IF;
  IF good_b THEN
    n_good := n_good + 1.0;
  END_IF;
  IF good_c THEN
    n_good := n_good + 1.0;
  END_IF;

  q_fail := n_good <= 0.0;

  (* Deviation monitor: any two good channels differ by more than dev_max (inline IF instead of ABS, library convention) *)
  q_dev := FALSE;
  IF dev_max > 0.0 THEN
    IF good_a AND good_b THEN
      IF (a - b > dev_max) OR (b - a > dev_max) THEN
        q_dev := TRUE;
      END_IF;
    END_IF;
    IF good_a AND good_c THEN
      IF (a - c > dev_max) OR (c - a > dev_max) THEN
        q_dev := TRUE;
      END_IF;
    END_IF;
    IF good_b AND good_c THEN
      IF (b - c > dev_max) OR (c - b > dev_max) THEN
        q_dev := TRUE;
      END_IF;
    END_IF;
  END_IF;

  IF n_good >= 3.0 THEN
    (* 3 good: take the median *)
    IF (a >= b AND a <= c) OR (a <= b AND a >= c) THEN
      out := a;
    ELSIF (b >= a AND b <= c) OR (b <= a AND b >= c) THEN
      out := b;
    ELSE
      out := c;
    END_IF;
  ELSIF n_good >= 2.0 THEN
    (* 2 good: take the average *)
    IF NOT good_a THEN
      out := (b + c) / 2.0;
    ELSIF NOT good_b THEN
      out := (a + c) / 2.0;
    ELSE
      out := (a + b) / 2.0;
    END_IF;
  ELSIF n_good >= 1.0 THEN
    (* 1 good: pass-through *)
    IF good_a THEN
      out := a;
    ELSIF good_b THEN
      out := b;
    ELSE
      out := c;
    END_IF;
  END_IF;
  (* 0 good: out holds the previous scan's value, q_fail signals it *)
END_FUNCTION_BLOCK

(* ---- fb_motor.st ---- *)
(*
  FB_MOTOR — motor start/stop control, with run-feedback monitoring and fault latch.

  Purpose: standard start/stop wrapper for single-speed motors such as belt conveyors,
  fans and pumps.
  Example: in remote mode an HMI/supervisory start/stop command -> contactor output,
  and a timed mismatch of the run feedback (contactor aux contact / current relay)
  faults the motor to stop.

  Behavior:
    1) Fault monitoring: a mismatch between out_run and run_fb persisting for
       fb_timeout_s (manual dt_s accumulation) -> fault latched; an external fault
       fault_in (thermal overload / drive fault, etc.) -> fault. reset with fault_in
       already cleared clears the latch.
    2) Command latch: cmd_start (level or momentary) sets out_run when remote and
       fault-free; cmd_stop or fault resets it (stop takes priority).
    3) Status word status: 0 stopped, 1 starting (output on, feedback not yet seen),
       2 running, 3 faulted.

  Inputs:
    cmd_start    BOOL  start command
    cmd_stop     BOOL  stop command (priority)
    remote       BOOL  remote permissive (gates start only; does not force a stop)
    run_fb       BOOL  run feedback
    fault_in     BOOL  external fault input
    reset        BOOL  fault reset
    fb_timeout_s REAL  feedback-mismatch tolerance time s
    dt_s         REAL  sample period s
  Outputs:
    out_run BOOL  run output (contactor / drive start)
    fault   BOOL  fault (latched)
    status  INT   0 stopped / 1 starting / 2 running / 3 faulted
*)
FUNCTION_BLOCK FB_MOTOR
  VAR_INPUT
    cmd_start    : BOOL;
    cmd_stop     : BOOL;
    remote       : BOOL := TRUE;
    run_fb       : BOOL;
    fault_in     : BOOL;
    reset        : BOOL;
    fb_timeout_s : REAL := 5.0;
    dt_s         : REAL := 0.1;
  END_VAR
  VAR_OUTPUT
    out_run : BOOL;
    fault   : BOOL;
    status  : INT;
  END_VAR
  VAR
    mism_t : REAL; (* feedback-mismatch accumulated time s *)
  END_VAR

  (* 1) Fault monitoring *)
  IF out_run <> run_fb THEN
    mism_t := mism_t + dt_s;
  ELSE
    mism_t := 0.0;
  END_IF;
  IF fb_timeout_s > 0.0 AND mism_t >= fb_timeout_s THEN
    fault := TRUE;
  END_IF;
  IF fault_in THEN
    fault := TRUE;
  END_IF;
  IF reset AND NOT fault_in THEN
    fault  := FALSE;
    mism_t := 0.0;
  END_IF;

  (* 2) Command latch (stop/fault priority) *)
  IF cmd_start AND remote AND NOT fault THEN
    out_run := TRUE;
  END_IF;
  IF cmd_stop OR fault THEN
    out_run := FALSE;
  END_IF;

  (* 3) Status word *)
  IF fault THEN
    status := 3;
  ELSIF out_run AND run_fb THEN
    status := 2;
  ELSIF out_run THEN
    status := 1;
  ELSE
    status := 0;
  END_IF;
END_FUNCTION_BLOCK

(* ---- fb_motor_rev.st ---- *)
(*
  FB_MOTOR_REV — bidirectional (forward/reverse) motor control, with reversal interlock,
  run-feedback monitoring and fault latch.

  ~ Standard reversing-motor block (reversing motor / forward-reverse starter, including
  the reversal-interlock delay), found in every major DCS/PLC standard library.

  Purpose: standard wrapper for reversible-running equipment such as agitators, hoists,
  bidirectional conveyors and gate-opening motors (pattern following FB_MOTOR: command
  latch + feedback-timeout fault latch).

  Behavior:
    1) Fault monitoring: fb_fwd and fb_rev TRUE at once -> feedback/contactor fault,
       immediate fault; an output-feedback mismatch (q_fwd<>fb_fwd or q_rev<>fb_rev)
       persisting for fb_timeout_s (manual dt_s accumulation) -> fault. All latched;
       cleared by reset with the dual-feedback condition cleared.
    2) Direction command latch (stop/fault priority): cmd_fwd / cmd_rev set the
       corresponding direction request (a both-direction command in the same scan is
       treated as a conflict, no action); stop or fault clears all requests.
    3) Reversal interlock: on a reversal (the reverse request is still present, or the
       reverse feedback is still turning), both outputs are forced fully stopped, and a
       new-direction output is allowed only after reversal_delay_s -- the contactor
       arc-quench / mechanical run-down time. reversal_delay_s should be less than
       fb_timeout_s (residual feedback rotation during the interlock wait is covered by
       the timeout tolerance).
    4) Status word state: 0 stopped / 1 forward / 2 reverse / 3 faulted / 4 reversal wait.

  Inputs:
    cmd_fwd          BOOL  forward command
    cmd_rev          BOOL  reverse command
    stop             BOOL  stop command (priority)
    fb_fwd           BOOL  forward run feedback
    fb_rev           BOOL  reverse run feedback
    fb_timeout_s     REAL  feedback-mismatch tolerance time s
    reversal_delay_s REAL  reversal full-stop interlock time s
    reset            BOOL  fault reset
    dt_s             REAL  sample period s
  Outputs:
    q_fwd BOOL  forward output
    q_rev BOOL  reverse output
    fault BOOL  fault (latched)
    state REAL  0 stopped / 1 forward / 2 reverse / 3 faulted / 4 reversal wait
*)
FUNCTION_BLOCK FB_MOTOR_REV
  VAR_INPUT
    cmd_fwd          : BOOL;
    cmd_rev          : BOOL;
    stop             : BOOL;
    fb_fwd           : BOOL;
    fb_rev           : BOOL;
    fb_timeout_s     : REAL := 5.0;
    reversal_delay_s : REAL := 2.0;
    reset            : BOOL;
    dt_s             : REAL := 0.1;
  END_VAR
  VAR_OUTPUT
    q_fwd : BOOL;
    q_rev : BOOL;
    fault : BOOL;
    state : REAL;
  END_VAR
  VAR
    want_fwd : BOOL; (* latched direction request *)
    want_rev : BOOL;
    wait_t   : REAL; (* reversal-interlock remaining time s *)
    mism_t   : REAL; (* feedback-mismatch accumulated time s *)
    conflict : BOOL; (* both-direction command in the same scan *)
  END_VAR

  (* 1) Fault monitoring *)
  IF fb_fwd AND fb_rev THEN
    fault := TRUE; (* both feedbacks active at once: welded contactor / feedback-circuit fault *)
  END_IF;
  IF (q_fwd <> fb_fwd) OR (q_rev <> fb_rev) THEN
    mism_t := mism_t + dt_s;
  ELSE
    mism_t := 0.0;
  END_IF;
  IF fb_timeout_s > 0.0 AND mism_t >= fb_timeout_s THEN
    fault := TRUE;
  END_IF;
  IF reset AND NOT (fb_fwd AND fb_rev) THEN
    fault  := FALSE;
    mism_t := 0.0;
  END_IF;

  (* 2) Direction command latch (stop/fault priority; a both-direction command in the same scan conflicts, no action) *)
  conflict := cmd_fwd AND cmd_rev;
  IF cmd_fwd AND NOT conflict AND NOT fault AND NOT stop THEN
    IF want_rev OR fb_rev THEN
      wait_t := reversal_delay_s; (* reverse still commanded / still turning: full-stop interlock first *)
    END_IF;
    want_fwd := TRUE;
    want_rev := FALSE;
  ELSIF cmd_rev AND NOT conflict AND NOT fault AND NOT stop THEN
    IF want_fwd OR fb_fwd THEN
      wait_t := reversal_delay_s;
    END_IF;
    want_rev := TRUE;
    want_fwd := FALSE;
  END_IF;
  IF stop OR fault THEN
    want_fwd := FALSE;
    want_rev := FALSE;
  END_IF;

  (* 3) Reversal-interlock timing (manual dt_s decrement) *)
  IF wait_t > 0.0 THEN
    wait_t := wait_t - dt_s;
    IF wait_t < 0.0 THEN
      wait_t := 0.0;
    END_IF;
  END_IF;

  (* 4) Output: during the interlock both outputs are forced fully stopped *)
  q_fwd := want_fwd AND wait_t <= 0.0;
  q_rev := want_rev AND wait_t <= 0.0;

  (* 5) Status word *)
  IF fault THEN
    state := 3.0;
  ELSIF wait_t > 0.0 AND (want_fwd OR want_rev) THEN
    state := 4.0;
  ELSIF q_fwd THEN
    state := 1.0;
  ELSIF q_rev THEN
    state := 2.0;
  ELSE
    state := 0.0;
  END_IF;
END_FUNCTION_BLOCK

(* ---- fb_mov.st ---- *)
(*
  FB_MOV — motor-operated valve (open/stop/close three commands + ZSO/ZSC dual limits + travel timeout).

  ~ Standard motor-operated-valve block (open/stop/close type, with travel monitoring),
  found in every major DCS/PLC standard library.

  Purpose: standard wrapper for "open-stop-close"-type motor-operated valves such as
  motorized gate/butterfly valves. Difference from FB_VALVE (two-position valve, single
  held output): this block is dual-direction pulse-driven with mid-travel stop, and the
  motor stops automatically at the limit; difference from FB_PID_3STEP (modulating step
  type): this block does only full-open/full-close/mid-stop sequential operations, no
  closed-loop control.

  Behavior:
    1) Fault monitoring: zso and zsc TRUE at once -> limit-switch fault, immediate fault;
       travel (an output active in either direction and the target limit not reached)
       exceeding travel_s -> travel-timeout fault (stuck valve / lost limit), and the
       outputs stop. All latched; cleared by reset with the dual-limit condition cleared
       (the travel timer is cleared in step).
    2) Commands: cmd_stop or fault -> both outputs stop (priority; cmd_open and cmd_close
       commanded together in the same scan is treated as a conflict, handled as stop);
       cmd_open latches the open output, cmd_close latches the close output (mutually
       exclusive, a new command is a new travel, the travel timer is cleared).
    3) Stop-at-position: zso reached during q_open -> stop the open output; zsc reached
       during q_close -> stop the close output.
    4) Status word pos_state: 0 fully closed / 1 opening / 2 fully open / 3 closing /
       4 faulted; a mid-stop (no output and not at a limit) holds the previous status value.

  Inputs:
    cmd_open  BOOL  open command
    cmd_close BOOL  close command
    cmd_stop  BOOL  stop command (priority, mid-stop)
    zso       BOOL  open limit
    zsc       BOOL  close limit
    travel_s  REAL  travel timeout s (<= 0 = not monitored)
    reset     BOOL  fault reset
    dt_s      REAL  sample period s
  Outputs:
    q_open    BOOL  open-direction output
    q_close   BOOL  close-direction output
    pos_state REAL  0 fully closed / 1 opening / 2 fully open / 3 closing / 4 faulted
    fault     BOOL  fault (latched)
*)
FUNCTION_BLOCK FB_MOV
  VAR_INPUT
    cmd_open  : BOOL;
    cmd_close : BOOL;
    cmd_stop  : BOOL;
    zso       : BOOL;
    zsc       : BOOL;
    travel_s  : REAL := 60.0;
    reset     : BOOL;
    dt_s      : REAL := 0.1;
  END_VAR
  VAR_OUTPUT
    q_open    : BOOL;
    q_close   : BOOL;
    pos_state : REAL;
    fault     : BOOL;
  END_VAR
  VAR
    travel_t : REAL; (* current-travel accumulated time s *)
  END_VAR

  (* 1) Dual-limit fault (immediate) *)
  IF zso AND zsc THEN
    fault := TRUE; (* both limits active at once: limit-switch fault *)
  END_IF;

  (* Reset (no effect while the dual-limit condition is still present) *)
  IF reset AND NOT (zso AND zsc) THEN
    fault    := FALSE;
    travel_t := 0.0;
  END_IF;

  (* 2) Command latch: stop/fault/both-commands-same-scan -> full stop; open and close mutually exclusive, a new command is a new travel *)
  IF cmd_stop OR fault OR (cmd_open AND cmd_close) THEN
    q_open  := FALSE;
    q_close := FALSE;
  ELSIF cmd_open THEN
    IF NOT q_open THEN
      travel_t := 0.0; (* new travel: clear the timer *)
    END_IF;
    q_open  := TRUE;
    q_close := FALSE;
  ELSIF cmd_close THEN
    IF NOT q_close THEN
      travel_t := 0.0;
    END_IF;
    q_close := TRUE;
    q_open  := FALSE;
  END_IF;

  (* 3) Stop-at-position *)
  IF q_open AND zso THEN
    q_open := FALSE;
  END_IF;
  IF q_close AND zsc THEN
    q_close := FALSE;
  END_IF;

  (* 4) Travel timeout (manual dt_s accumulation) *)
  IF q_open OR q_close THEN
    travel_t := travel_t + dt_s;
    IF travel_s > 0.0 AND travel_t >= travel_s THEN
      fault   := TRUE; (* travel timeout: stuck valve / lost limit *)
      q_open  := FALSE;
      q_close := FALSE;
    END_IF;
  ELSE
    travel_t := 0.0;
  END_IF;

  (* 5) Status word (a mid-stop holds the previous status value) *)
  IF fault THEN
    pos_state := 4.0;
  ELSIF zso THEN
    pos_state := 2.0;
  ELSIF zsc THEN
    pos_state := 0.0;
  ELSIF q_open THEN
    pos_state := 1.0;
  ELSIF q_close THEN
    pos_state := 3.0;
  END_IF;
END_FUNCTION_BLOCK

(* ---- fb_pid.st ---- *)
(*
  FB_PID — incremental (velocity-form) PID controller with anti-windup,
  bumpless transfer, feedforward, output tracking and setpoint ramp.

  ~ Universal PID essentials: SP ramp / output tracking / feedforward / auto-manual
    bumpless transfer (every major DCS/PLC standard library has an equivalent block).

  Typical use: a flow PID driving a variable-speed pump, direct-acting, where the
  output limits are the drive min/max frequency (e.g. 10..45 Hz — flow is pv, the
  drive frequency reference is out: out_min:=10.0, out_max:=45.0, direct := TRUE
  direct-acting — rising pv raises output).

  Algorithm (incremental + feedforward):
    sp_int := sp through an sp_rate-limited ramp (sp_rate <= 0 takes sp directly; first-scan alignment)
    e      := sp_int - pv (reverse-acting, default); direct=TRUE gives e := pv - sp_int
    dpid   := kp*(e - e_prev)                            -- proportional increment
            + kp*dt_s/ti_s * e (when ti_s>0)             -- integral increment
            + kp*td_s/dt_s * (e - 2*e_prev + e_prev2) (when td_s>0) -- derivative increment
    acc    := acc + dpid; out := acc + ff, clamped to [out_min, out_max]
    wrap-up  acc := out - ff (back-calculation)
  Anti-windup: output clamp + back-calculation + conditional integration (when the
  output is already at a limit and the integral increment keeps pushing toward that
  limit, the integral term is dropped).
  Mode priority: track (output tracking, for interlock forcing / external takeover)
  > NOT auto (manual) > auto. In track/manual the output follows the supplied value
  (clamped), the error history keeps updating, and returning to auto is bumpless.
  ff adds directly onto the pre-clamp output (feedforward takes effect immediately;
  back-calculation keeps ff changes, clamping and mode switching all bumpless).
  Backward compatible: the added inputs (ff/track/track_value/sp_rate) all have
  defaults, and at their defaults behavior is scan-for-scan identical to the old
  version, so existing calls need no changes; the added output dev does not affect
  legacy wiring.

  Inputs:
    pv          REAL  process value
    sp          REAL  setpoint
    kp          REAL  proportional gain
    ti_s        REAL  integral time s (0 = integral off)
    td_s        REAL  derivative time s (0 = derivative off, derivative term unfiltered)
    dt_s        REAL  sample period s (<=0 holds this scan, no action)
    direct      BOOL  TRUE = direct-acting (pv up -> out up), FALSE = reverse-acting
    auto        BOOL  TRUE auto / FALSE manual
    manual_out  REAL  manual output value
    out_min     REAL  output low limit (assumes out_min < out_max)
    out_max     REAL  output high limit
    ff          REAL  feedforward (added to output before clamp; feed via FB_LEADLAG for dynamic shaping)
    track       BOOL  output-tracking enable (highest priority, overrides auto/manual)
    track_value REAL  tracking value
    sp_rate     REAL  setpoint ramp rate limit units/s (0 = no rate limit)
  Outputs:
    out         REAL  control output (clamped in every mode)
    dev         REAL  deviation pv - sp_int (actual working deviation after the SP ramp)
*)
FUNCTION_BLOCK FB_PID
  VAR_INPUT
    pv          : REAL;
    sp          : REAL;
    kp          : REAL := 1.0;
    ti_s        : REAL := 0.0;
    td_s        : REAL := 0.0;
    dt_s        : REAL := 0.1;
    direct      : BOOL := FALSE;
    auto        : BOOL := TRUE;
    manual_out  : REAL := 0.0;
    out_min     : REAL := 0.0;
    out_max     : REAL := 100.0;
    ff          : REAL := 0.0;
    track       : BOOL := FALSE;
    track_value : REAL := 0.0;
    sp_rate     : REAL := 0.0;
  END_VAR
  VAR_OUTPUT
    out : REAL;
    dev : REAL;
  END_VAR
  VAR
    sp_int    : REAL; (* internal working setpoint after the ramp *)
    acc       : REAL; (* PID accumulator (excludes ff) *)
    e         : REAL;
    e_prev    : REAL;
    e_prev2   : REAL;
    p_term    : REAL;
    i_term    : REAL;
    d_term    : REAL;
    sp_step   : REAL;
    sp_delta  : REAL;
    init_done : BOOL; (* sp_int first-scan alignment flag *)
  END_VAR

  IF dt_s <= 0.0 THEN
    RETURN; (* invalid sample period: hold output and history unchanged *)
  END_IF;

  (* Setpoint ramp: when sp_rate > 0, sp_int approaches sp at the rate limit; first scan aligns directly *)
  IF NOT init_done THEN
    sp_int := sp;
    init_done := TRUE;
  ELSIF sp_rate > 0.0 THEN
    sp_step := sp_rate * dt_s;
    sp_delta := sp - sp_int;
    IF sp_delta > sp_step THEN
      sp_int := sp_int + sp_step;
    ELSIF sp_delta < 0.0 - sp_step THEN
      sp_int := sp_int - sp_step;
    ELSE
      sp_int := sp;
    END_IF;
  ELSE
    sp_int := sp;
  END_IF;

  dev := pv - sp_int;

  (* Control deviation; direct-acting flips the sign *)
  IF direct THEN
    e := pv - sp_int;
  ELSE
    e := sp_int - pv;
  END_IF;

  IF track THEN
    (* Output tracking: follows track_value unconditionally (interlock forcing / override takeover), highest priority *)
    out := track_value;
  ELSIF NOT auto THEN
    (* Manual: follows manual_out; the incremental form makes the return to auto naturally bumpless *)
    out := manual_out;
  ELSE
    p_term := kp * (e - e_prev);

    i_term := 0.0;
    IF ti_s > 0.0 THEN
      i_term := kp * dt_s / ti_s * e;
      (* Conditional integration: when the output is saturated and the integral still pushes toward the limit, drop the integral term this scan *)
      IF (out >= out_max AND i_term > 0.0) OR (out <= out_min AND i_term < 0.0) THEN
        i_term := 0.0;
      END_IF;
    END_IF;

    d_term := 0.0;
    IF td_s > 0.0 THEN
      d_term := kp * td_s / dt_s * (e - 2.0 * e_prev + e_prev2);
    END_IF;

    acc := acc + p_term + i_term + d_term;
    out := acc + ff; (* feedforward added before clamp *)
  END_IF;

  (* Output clamp (in the incremental form this also provides anti-windup) *)
  IF out > out_max THEN
    out := out_max;
  ELSIF out < out_min THEN
    out := out_min;
  END_IF;

  (* Back-calculation: acc always = clamped output - feedforward -> clamping / ff changes / manual / tracking all bumpless *)
  acc := out - ff;

  e_prev2 := e_prev;
  e_prev  := e;
END_FUNCTION_BLOCK
